(* IEC 61131-3 sources: plc-repo-template/tests/POUs/FB_Example_Test, 12 files *)

(* ---- FB_Example_Test.decl.st ---- *)
// Назначение: набор тестов CfUnit (coUnit 1.2.0.0) для FB_Example — включение и отключение
//             по порогам гистерезиса и на самих порогах, удержание состояния в зоне
//             гистерезиса, защёлка отказа измерения и квитирование, режимы Manual, Local,
//             OutOfService, режим по умолчанию, ограничение параметров, счётчик включений
//             и сброс через I_Resettable. Каждый тест работает со своим экземпляром FB_Example
//             (локальная переменная метода) и укладывается в один цикл.
// Автор:      kr0nsch
// Версия:     0.1.0
// Документ:   docs/TEST_REPORT.md
FUNCTION_BLOCK FB_Example_Test EXTENDS coUnit.FB_TestSuite
VAR CONSTANT
    // Уставка отключения и гистерезис: включение при значении <= 50 %, отключение при >= 60 %
    R_SP_PCT : REAL := 60.0;
    R_HYST_PCT : REAL := 10.0;
    R_ON_THRESHOLD_PCT : REAL := 50.0;  // порог включения: R_SP_PCT - R_HYST_PCT
    R_LOW_PCT : REAL := 40.0;           // ниже порога включения
    R_BAND_PCT : REAL := 55.0;          // внутри зоны гистерезиса
    R_HIGH_PCT : REAL := 70.0;          // выше уставки отключения
    // Параметры вне допустимых диапазонов GVL_Const
    R_SP_TOO_HIGH_PCT : REAL := 150.0;
    R_HYST_TOO_LOW_PCT : REAL := 0.1;
    // F_Clamp возвращает одну из своих границ без арифметики — сравнение точное
    R_DELTA : REAL := 0.0;
    UDI_TWO_SWITCH_ONS : UDINT := 2;    // ожидаемое число включений в тесте счётчика
END_VAR

(* ---- AcknowledgeClearsFaultWhenValid.method.decl.st ---- *)
// Квитирование при достоверном измерении снимает отказ, выход снова управляется.
METHOD PRIVATE AcknowledgeClearsFaultWhenValid
VAR
    fbDut : FB_Example;         // проверяемый экземпляр, новый при каждом вызове метода
    xAckResult : BOOL;          // результат Acknowledge()
END_VAR

(* ---- AcknowledgeKeepsFaultWhileInvalid.method.decl.st ---- *)
// Квитирование при недостоверном измерении отказ не снимает.
METHOD PRIVATE AcknowledgeKeepsFaultWhileInvalid
VAR
    fbDut : FB_Example;         // проверяемый экземпляр, новый при каждом вызове метода
    xAckResult : BOOL;          // результат Acknowledge()
END_VAR

(* ---- AutoHoldsStateInsideHysteresis.method.decl.st ---- *)
// Авторежим: внутри зоны гистерезиса выход сохраняет прежнее состояние в обе стороны.
METHOD PRIVATE AutoHoldsStateInsideHysteresis
VAR
    fbDut : FB_Example;         // проверяемый экземпляр, новый при каждом вызове метода
END_VAR

(* ---- AutoSwitchesOnBelowThreshold.method.decl.st ---- *)
// Авторежим: значение ниже порога включения (уставка - гистерезис) включает выход.
METHOD PRIVATE AutoSwitchesOnBelowThreshold
VAR
    fbDut : FB_Example;         // проверяемый экземпляр, новый при каждом вызове метода
END_VAR

(* ---- AutoThresholdsAreInclusive.method.decl.st ---- *)
// Авторежим: на пороге включения выход включается, на уставке — отключается.
METHOD PRIVATE AutoThresholdsAreInclusive
VAR
    fbDut : FB_Example;         // проверяемый экземпляр, новый при каждом вызове метода
END_VAR

(* ---- CountsSwitchOnsAndResetClears.method.decl.st ---- *)
// Счётчик считает включения по фронту выхода; Reset() через I_Resettable отключает
// выход и обнуляет счётчик.
METHOD PRIVATE CountsSwitchOnsAndResetClears
VAR
    fbDut : FB_Example;         // проверяемый экземпляр, новый при каждом вызове метода
    itfDut : I_Resettable;      // сброс через интерфейс, как в PRG_Main
    xResetResult : BOOL;        // результат Reset()
END_VAR

(* ---- DefaultModeIsOutOfService.method.decl.st ---- *)
// Пока режим не назначен (значение входа по умолчанию), выход отключён.
METHOD PRIVATE DefaultModeIsOutOfService
VAR
    fbDut : FB_Example;         // проверяемый экземпляр, новый при каждом вызове метода
END_VAR

(* ---- InvalidValueLatchesFault.method.decl.st ---- *)
// Отказ измерения в авторежиме: выход отключается, отказ держится и после
// восстановления измерения — до квитирования.
METHOD PRIVATE InvalidValueLatchesFault
VAR
    fbDut : FB_Example;         // проверяемый экземпляр, новый при каждом вызове метода
END_VAR

(* ---- LocalAndOutOfServiceSwitchOff.method.decl.st ---- *)
// Режимы Local и OutOfService снимают команду ПЛК при любом измерении и команде.
METHOD PRIVATE LocalAndOutOfServiceSwitchOff
VAR
    fbDut : FB_Example;         // проверяемый экземпляр, новый при каждом вызове метода
END_VAR

(* ---- ManualFollowsCommand.method.decl.st ---- *)
// Ручной режим: выход повторяет команду оператора, измерение на выход не влияет
// и отказ не фиксируется (docs/ASSUMPTIONS.md, C5).
METHOD PRIVATE ManualFollowsCommand
VAR
    fbDut : FB_Example;         // проверяемый экземпляр, новый при каждом вызове метода
END_VAR

(* ---- ParametersAreClamped.method.decl.st ---- *)
// Уставка и гистерезис вне допустимых диапазонов ограничиваются границами из GVL_Const.
METHOD PRIVATE ParametersAreClamped
VAR
    fbDut : FB_Example;         // проверяемый экземпляр, новый при каждом вызове метода
END_VAR
